DEVICE_TYPE TestDevice (* Device type for the import export system *)
  (* Standard: 61499-1; Description: Copyright (c) 2026 Martin Erich Jobst This program and the accompanying materials are made available under the terms of the Eclipse Public License 2.0 which is available at https://www.eclipse.org/legal/epl-2.0/ SPDX-License-Identifier: EPL-2.0 *)
  (* Version 1.0, 2026-10-23, Martin Jobst *)
  {SET_ATTRIBUTE(IntegerAttribute, 12)}
  VAR_INPUT
    DEVICE_ID : DINT := DINT#1;
  END_VAR
  RESOURCE LocalResource : TestResource(RESOURCE_ID := DINT#3) (* Fixture resource *)
    {SET_ATTRIBUTE(IntegerAttribute, 11)}
  END_RESOURCE
END_DEVICE_TYPE
